(* IEC 61131-3 sources: plcassist-cli/packages/volt-lsp-iec/test-corpus/awa-palletizer/Device/Plc Logic/Application/Library Manager/CAA Mathematics, 39 files *)

(* ---- GLOBALCONSTANTS.gvl ---- *)
VAR_GLOBAL
	PI : LREAL := 3.1415926535897931;
END_VAR

(* ---- VERSIONCONSTANTS.gvl ---- *)
VAR_GLOBAL
	GC_BYVERSION : BYTE := 1;
	GC_VERSION_1 : BYTE := 0;
END_VAR

(* ---- ADDMULTIPLICATEDVECTOR.fun ---- *)
FUNCTION ADDMULTIPLICATEDVECTOR : BOOL
VAR_INPUT
	PV1 : POINTER TO Vector3d;
	PV2 : POINTER TO Vector3d;
	LRFACTOR : LREAL;
	PV : POINTER TO Vector3D;
END_VAR
END_FUNCTION

(* ---- ATAN2.fun ---- *)
FUNCTION ATAN2 : LREAL
VAR_INPUT
	LRSINUS : LREAL;
	LRCOSINUS : LREAL;
END_VAR
END_FUNCTION

(* ---- ATAN2_FUNC.fun ---- *)
FUNCTION ATAN2_FUNC : LREAL
VAR_INPUT
	LRSINUS : LREAL;
	LRCOSINUS : LREAL;
END_VAR
END_FUNCTION

(* ---- FMOD.fun ---- *)
FUNCTION FMOD : LREAL
VAR_INPUT
	LRX : LREAL;
	LRM : LREAL;
END_VAR
END_FUNCTION

(* ---- GETLIBVERSION.fun ---- *)
FUNCTION GETLIBVERSION : VERSION
END_FUNCTION

(* ---- GETLIBVERSIONNUMBER.fun ---- *)
FUNCTION GETLIBVERSIONNUMBER : DWORD
END_FUNCTION

(* ---- GETSUPPLIERVERSION.fun ---- *)
FUNCTION GETSUPPLIERVERSION : WORD
VAR_INPUT
	XDUMMY : BOOL;
END_VAR
END_FUNCTION

(* ---- ISLIBRELEASED.fun ---- *)
FUNCTION ISLIBRELEASED : BOOL
END_FUNCTION

(* ---- MAKENORMED3D.fun ---- *)
FUNCTION MAKENORMED3D : BOOL
VAR_INPUT
	PV : POINTER TO VECTOR3D;
END_VAR
END_FUNCTION

(* ---- NORM3D.fun ---- *)
FUNCTION NORM3D : LREAL
VAR_INPUT
	PV : POINTER TO VECTOR3D;
END_VAR
END_FUNCTION

(* ---- POLYNOMIALVALUE.fun ---- *)
FUNCTION POLYNOMIALVALUE : LREAL
VAR_INPUT
	SIDEGREE : SINT;
	PLR : POINTER TO LREAL;
	LRVALUE : LREAL;
END_VAR
END_FUNCTION

(* ---- PROJECTPOINTONLINE.fun ---- *)
FUNCTION PROJECTPOINTONLINE : BOOL
VAR_INPUT
	PLINE : POINTER TO LINE_3D;
	PVORIG : POINTER TO Vector3D;
	PVPROJ : POINTER TO Vector3D;
END_VAR
END_FUNCTION

(* ---- PROJECTPOINTONPLANE.fun ---- *)
FUNCTION PROJECTPOINTONPLANE : LREAL
VAR_INPUT
	PPLANE : POINTER TO Plane_H;
	PVORIG : POINTER TO VECTOR3D;
	PVPROJ : POINTER TO VECTOR3D;
END_VAR
END_FUNCTION

(* ---- SCALPROD3D.fun ---- *)
FUNCTION SCALPROD3D : LREAL
VAR_INPUT
	PV1 : POINTER TO Vector3d;
	PV2 : POINTER TO Vector3d;
END_VAR
END_FUNCTION

(* ---- SCALPROD3DSTAND.fun ---- *)
FUNCTION SCALPROD3DSTAND : LREAL
VAR_INPUT
	PV1 : POINTER TO Vector3d;
	PV2 : POINTER TO Vector3d;
END_VAR
END_FUNCTION

(* ---- SGN.fun ---- *)
FUNCTION SGN : INT
VAR_INPUT
	LR : LREAL;
END_VAR
END_FUNCTION

(* ---- SUBVECTOR.fun ---- *)
FUNCTION SUBVECTOR : BOOL
VAR_INPUT
	PV1 : POINTER TO Vector3d;
	PV2 : POINTER TO Vector3d;
	PV : POINTER TO Vector3D;
END_VAR
END_FUNCTION

(* ---- CALCHESSEREPRESENTATION.fb ---- *)
FUNCTION_BLOCK CALCHESSEREPRESENTATION
VAR_INPUT
	VP1 : POINTER TO Vector3D;
	VP2 : POINTER TO Vector3D;
	VP3 : POINTER TO Vector3D;
END_VAR
VAR_OUTPUT
	PLANE : PLANE_H;
	XERROR : BOOL;
END_VAR
VAR
	V1 : Vector3D;
	V2 : Vector3D;
	VN : Vector3D;
	CP : CrossProductNormed;
END_VAR
END_FUNCTION_BLOCK

(* ---- CALCROOTLIN.fb ---- *)
FUNCTION_BLOCK CALCROOTLIN
VAR_INPUT
	LRPARAM1 : LREAL;
	LRPARAM0 : LREAL;
END_VAR
VAR_OUTPUT
	BYROOTS : BYTE;
	LRROOT : LREAL;
END_VAR
END_FUNCTION_BLOCK

(* ---- CALCROOTPARABLE.fb ---- *)
FUNCTION_BLOCK CALCROOTPARABLE
VAR_INPUT
	LRPARAM2 : LREAL;
	LRPARAM1 : LREAL;
	LRPARAM0 : LREAL;
END_VAR
VAR_OUTPUT
	BYROOTS : BYTE;
	LRROOT0 : LREAL;
	LRROOT1 : LREAL;
END_VAR
VAR
	D : LREAL;
END_VAR
END_FUNCTION_BLOCK

(* ---- CARTESIANTOPOLAR.fb ---- *)
FUNCTION_BLOCK CARTESIANTOPOLAR
VAR_INPUT
	LRX : LREAL;
	LRY : LREAL;
END_VAR
VAR_OUTPUT
	LRANGLE : LREAL;
	LRDISTANCE : LREAL;
END_VAR
END_FUNCTION_BLOCK

(* ---- CHARCURVE_DINT.fb ---- *)
FUNCTION_BLOCK CHARCURVE_DINT
VAR_INPUT
	DIINPUTVALUE : DINT;
	USINOPOINTS : USINT;
END_VAR
VAR_OUTPUT
	DIOUTPUTVALUE : DINT;
	XERROR : BOOL;
	WERRORID : WORD;
END_VAR
VAR_IN_OUT
	AP2DIPOINTS : ARRAY [0..10] OF POINT2_DINT;
END_VAR
VAR
	I : INT;
END_VAR
END_FUNCTION_BLOCK

(* ---- CHARCURVE_LREAL.fb ---- *)
FUNCTION_BLOCK CHARCURVE_LREAL
VAR_INPUT
	LRINPUTVALUE : LREAL;
	USINOPOINTS : USINT;
END_VAR
VAR_OUTPUT
	LROUTPUTVALUE : LREAL;
	XERROR : BOOL;
	WERRORID : WORD;
END_VAR
VAR_IN_OUT
	AP2LRPOINTS : ARRAY [0..10] OF POINT2_LREAL;
END_VAR
VAR
	I : INT;
END_VAR
END_FUNCTION_BLOCK

(* ---- CROSSPRODUCT.fb ---- *)
FUNCTION_BLOCK CROSSPRODUCT
VAR_INPUT
	V1 : Vector3d;
	V2 : Vector3d;
END_VAR
VAR_OUTPUT
	V : Vector3D;
END_VAR
END_FUNCTION_BLOCK

(* ---- CROSSPRODUCTNORMED.fb ---- *)
FUNCTION_BLOCK CROSSPRODUCTNORMED
VAR_INPUT
	V1 : Vector3d;
	V2 : Vector3d;
END_VAR
VAR_OUTPUT
	V : Vector3D;
	XERROR : BOOL;
END_VAR
VAR
	CP : CrossProduct;
END_VAR
END_FUNCTION_BLOCK

(* ---- DERIVATIVE.fb ---- *)
FUNCTION_BLOCK DERIVATIVE
VAR_INPUT
	XENABLE : BOOL;
	LRINPUTVALUE : LREAL;
	UDITM : UDINT;
END_VAR
VAR_OUTPUT
	LRDERIVATIVE : LREAL;
	XVALID : BOOL;
END_VAR
VAR
	LRX3 : LREAL;
	LRX2 : LREAL;
	LRX1 : LREAL;
	UDIT2 : UDINT;
	UDIT1 : UDINT;
	XOLDENABLE : BOOL;
	SI : SINT;
END_VAR
END_FUNCTION_BLOCK

(* ---- HYSTERESIS_DINT.fb ---- *)
FUNCTION_BLOCK HYSTERESIS_DINT
VAR_INPUT
	DIVALUE : DINT;
	DILIMITPOS : DINT;
	DILIMITNEG : DINT;
END_VAR
VAR_OUTPUT
	XOUT : BOOL;
END_VAR
END_FUNCTION_BLOCK

(* ---- HYSTERESIS_LREAL.fb ---- *)
FUNCTION_BLOCK HYSTERESIS_LREAL
VAR_INPUT
	LRVALUE : LREAL;
	LRLIMITPOS : LREAL;
	LRLIMITNEG : LREAL;
END_VAR
VAR_OUTPUT
	XOUT : BOOL;
END_VAR
END_FUNCTION_BLOCK

(* ---- INTEGRAL.fb ---- *)
FUNCTION_BLOCK INTEGRAL
VAR_INPUT
	XENABLE : BOOL;
	LRINPUTVALUE : LREAL;
	UDITM : UDINT;
END_VAR
VAR_OUTPUT
	LRINTEGRAL : LREAL;
	XOVERFLOW : BOOL := FALSE;
END_VAR
VAR
	XOLDENABLE : BOOL;
END_VAR
END_FUNCTION_BLOCK

(* ---- LIMITALARM_DINT.fb ---- *)
FUNCTION_BLOCK LIMITALARM_DINT
VAR_INPUT
	DIVALUE : DINT;
	DILIMITPOS : DINT;
	DILIMITNEG : DINT;
END_VAR
VAR_OUTPUT
	XEXCEEDSPOS : BOOL;
	XEXCEEDSNEG : BOOL;
	XINLIMITS : BOOL;
END_VAR
END_FUNCTION_BLOCK

(* ---- LIMITALARM_LREAL.fb ---- *)
FUNCTION_BLOCK LIMITALARM_LREAL
VAR_INPUT
	LRVALUE : LREAL;
	LRLIMITPOS : LREAL;
	LRLIMITNEG : LREAL;
END_VAR
VAR_OUTPUT
	XEXCEEDSPOS : BOOL;
	XEXCEEDSNEG : BOOL;
	XINLIMITS : BOOL;
END_VAR
END_FUNCTION_BLOCK

(* ---- LINEARTRAFO.fb ---- *)
FUNCTION_BLOCK LINEARTRAFO
VAR_INPUT
	LRINPUTVALUE : LREAL;
	LRINPUT1 : LREAL;
	LRINPUT2 : LREAL;
	LROUTPUT1 : LREAL;
	LROUTPUT2 : LREAL;
END_VAR
VAR_OUTPUT
	LROUTPUTVALUE : LREAL;
	XOUTOFLIMITS : BOOL;
END_VAR
VAR
	LRDIFF : LREAL;
END_VAR
END_FUNCTION_BLOCK

(* ---- MEASUREFREQUENCE.fb ---- *)
FUNCTION_BLOCK MEASUREFREQUENCE
VAR_INPUT
	XENABLE : BOOL;
	XINPUT : BOOL;
	USIPERIODS : USINT (1..10) := 1;
END_VAR
VAR_OUTPUT
	LRFREQUENCY : LREAL;
	XVALID : BOOL;
END_VAR
VAR
	TIMOLD : TIME;
	T2 : TIME;
	UDIDIFF : UDINT;
	AUDIDIFF : ARRAY [0..9] OF UDINT;
	IV : INT;
	IB : INT;
	I : INT;
	XOLDENABLE : BOOL;
	XOLDINPUT : BOOL;
	USIOLDPERIODS : USINT;
END_VAR
END_FUNCTION_BLOCK

(* ---- POLARTOCARTESIAN.fb ---- *)
FUNCTION_BLOCK POLARTOCARTESIAN
VAR_INPUT
	LRANGLE : LREAL;
	LRDISTANCE : LREAL;
END_VAR
VAR_OUTPUT
	LRX : LREAL;
	LRY : LREAL;
END_VAR
END_FUNCTION_BLOCK

(* ---- STATISTICS_DINT.fb ---- *)
FUNCTION_BLOCK STATISTICS_DINT
VAR_INPUT
	XENABLE : BOOL;
	DIINPUT : DINT;
END_VAR
VAR_OUTPUT
	DIMIN : DINT := 16#7FFFFFFF;
	DIMAX : DINT := DWORD_TO_DINT(16#80000000);
	DIAVERAGE : DINT;
	XOVERRUN : BOOL;
END_VAR
VAR
	DISUM : DINT;
	UDICOUNTER : UDINT;
	XOLDENABLE : BOOL;
END_VAR
END_FUNCTION_BLOCK

(* ---- STATISTICS_LREAL.fb ---- *)
FUNCTION_BLOCK STATISTICS_LREAL
VAR_INPUT
	XENABLE : BOOL;
	LRINPUT : LREAL;
END_VAR
VAR_OUTPUT
	LRMIN : LREAL := LREAL#1E+80;
	LRMAX : LREAL := LREAL#-1E+80;
	LRAVERAGE : LREAL;
	XOVERRUN : BOOL;
END_VAR
VAR
	UDICOUNTER : UDINT;
	LRSUM : LREAL;
	XOLDENABLE : BOOL;
END_VAR
END_FUNCTION_BLOCK

(* ---- VARIANCE.fb ---- *)
FUNCTION_BLOCK VARIANCE
VAR_INPUT
	XENABLE : BOOL;
	LRINPUTVALUE : LREAL;
END_VAR
VAR_OUTPUT
	LRVARIANCE : LREAL;
END_VAR
VAR
	UDIZ : UDINT;
	LRA : LREAL;
	LRB : LREAL;
END_VAR
END_FUNCTION_BLOCK
